RoboDK station: car_painting_cell_v1.rdk

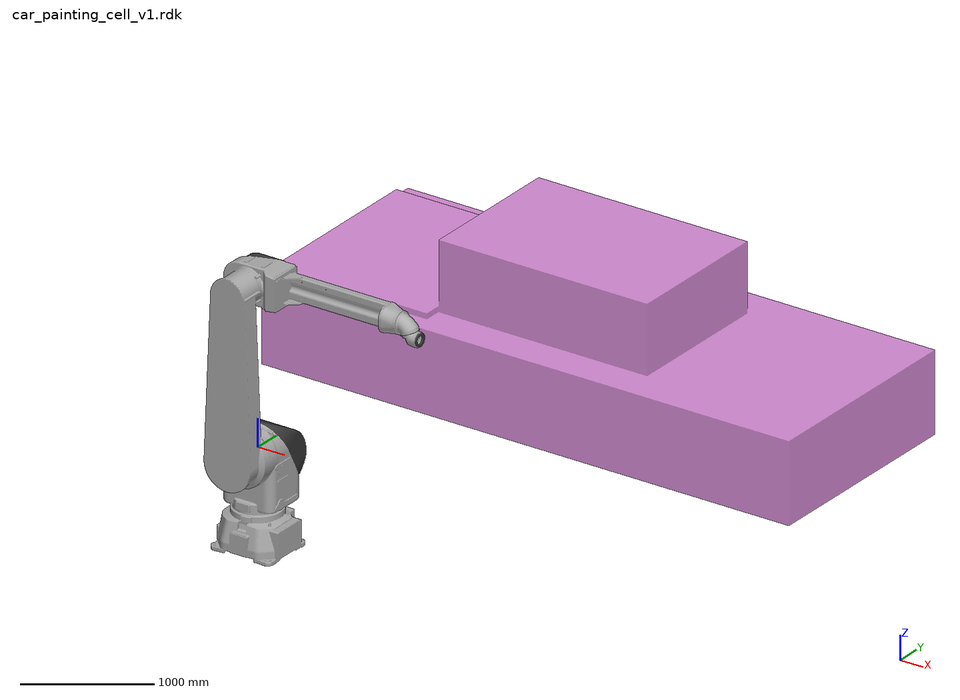
[picture v0: the station drawn from its stored meshes, robots at their saved joint values, targets as dots, program paths as lines]
Station car_painting_cell_v1 (saved by RoboDK 6.1.1). Poses are relative to the parent item; angles as X-Y-Z fixed-axis rotations.
  - frame Fanuc P-250iB RH Base at (0, 0, 820) mm
    - robot Fanuc P-250iB RH: 6 axes, payload 15 kg, reach 2800 mm, repeatability 0.07 mm, weight 530 kg
        modified DH rows (alpha deg, a mm, theta deg, d mm): 0, 0, 0, 820; -90, 0, -90, 0; 0, 1400, 0, 0; -90, 0, -90, 1362.687; 70, 0, 0, 106.416; -70, 0, 0, 81.885
        base shift (0, 0, -820) mm
        joint limits [-160, -45, -205, -360, -360, -360] to [160, 120, 165, 360, 360, 360]; home [0, 0, 0, 0, 0, 0]; saved at [0, 0, 0, 0, 0, 0]
  - object simple_car at (1000, 3000, 0) mm, size 4800 x 1900 x 1300 mm, geometry from simple_car.stl
